// TIA Portal V21 export
// export: Created 2026-11-11T00:47:18.0894613Z, ExportSetting WithDefaults, DisplayName Totally Integrated Automation Portal, DisplayVersion V21 Update 3, DisplayName STEP 7 Professional, DisplayVersion V21 Update 3, DisplayName STEP 7 Safety, DisplayVersion V21, DisplayName Tech WebApplication, DisplayVersion V21, DisplayName WinCC Basic/Comfort/Advanced, DisplayVersion V21 Update 3, DisplayName WinCC Unified, DisplayVersion V21 Update 3
FUNCTION_BLOCK "FB_Fbd_ex048"   // FB91, FBD
{ S7_Optimized_Access := 'TRUE' }
VERSION : 0.1
// stored: AutoNumber true, IsIECCheckEnabled false, IsRetainMemResEnabled false, MemoryReserve 100, SetENOAutomatically false, UDAEnableTagReadback false
   VAR_INPUT
      v_id : HW_SUBMODULE;
   END_VAR
   VAR_OUTPUT
      v_status : DWord;
   END_VAR
   VAR_IN_OUT
      v_outputs : Array[0..99] of Byte;
   END_VAR
   VAR
      inst { S7_SetPoint := 'True'} : SETIO;
   END_VAR
BEGIN

REGION Network 1: SETIO - Write all outputs of a submodule
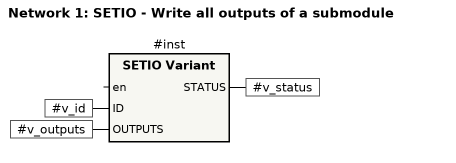
   #inst(ID := #v_id, OUTPUTS := #v_outputs, STATUS => #v_status);   // SETIO
END_REGION
END_FUNCTION_BLOCK
